(*
SPDX-FileCopyrightText: © 2026 Oleksandr Tiutyk <trofimich@gmail.com>
SPDX-License-Identifier: MIT
License: https://opensource.org/license/mit
*)

(*!
<summary>
Beckhoff EL3314: 4-channel thermocouple input terminal (J, K, T, E, N, R, S, B, C).
</summary>
<description>
Process image mapping structure for the EL3314 4-channel thermocouple input terminal.
When used for I/O, link located fields or their containing buffers to the matching selected PDOs.
The record is not a packed wire buffer; compiler padding is not part of the device specification.
Unlinked/default values do not prove valid I/O. The caller evaluates bus/channel validity before use.
Use one owner task per instance and externally synchronize other access; multi-field snapshots are not atomic.
Copies store data without creating hardware links. Keep borrowed field references valid while consumers are bound.
This passive record performs no validation, synchronization, configuration or protocol advancement.
Select standard status-plus-INT16 PDOs; compact layouts are unsupported. Configure presentation explicitly:
0.1/0.01 deg C per digit follows the device setting, not this record.
</description>
*)
TYPE EL3314 :
STRUCT
	Ch1 : THERMOCOUPLE_INPUT_CHANNEL;
	Ch2 : THERMOCOUPLE_INPUT_CHANNEL;
	Ch3 : THERMOCOUPLE_INPUT_CHANNEL;
	Ch4 : THERMOCOUPLE_INPUT_CHANNEL;
END_STRUCT
END_TYPE

(* stored: Version 1.1.0.1, ProductVersion 3.1.4026.20
   DUT EL3314: Id {1f765c08-8b95-4b50-b359-1f47d8cd9e76} *)
